// TIA Portal V20 export
Screen "170FX1Layout"  1276x673
  ScreenItem "Graphic view_1" at 215,132 size 858x332  Type=HmiGraphicView
  ScreenItem "Line_Header_X0_Y64" at 0,64 size 1276x0  Type=HmiLine
  ScreenItem "permanentareaborderrectangle" at 0,0 size 0x0  Type=HmiRectangle
  ScreenItem "Button_Back" at 2,2 size 90x60  Type=HmiButton
  ScreenItem "Move_Legend" at 1182,2 size 90x60  Type=HmiButton
  ScreenItem "Fusszeile_Button_ManualOPMode1_2" at 279,2 size 90x60  Type=HmiButton
  ScreenItem "文本域_3" at 1107,71 size 139x22  Type=HmiTextBox
  ScreenItem "LSicar_Valve8Pos_LeftHomeRightWork_WithPB_5" at 1099,95 size 160x53  Type=HmiFaceplateContainer
  ScreenItem "文本域_1" at 1107,160 size 156x23  Type=HmiTextBox
  ScreenItem "LSicar_Valve8Pos_LeftHomeRightWork_WithPB_1" at 1099,183 size 160x53  Type=HmiFaceplateContainer
  ScreenItem "文本域_22" at 1124,475 size 104x23  Type=HmiTextBox
  ScreenItem "面板容器_23" at 1171,508 size 96x32  Type=HmiFaceplateContainer
  ScreenItem "面板容器_22" at 1061,508 size 96x32  Type=HmiFaceplateContainer
  ScreenItem "面板容器_2" at 1087,4 size 88x58  Type=HmiFaceplateContainer
  ScreenItem "OPMode1_Blocked" at 1164,6 size 14x14  Type=HmiGraphicView
  ScreenItem "OPMode4_Foreground_Blocked" at 1088,4 size 88x58  Type=HmiGraphicView
  ScreenItem "Fusszeile_Button_ManualOPMode1_1" at 95,2 size 90x60  Type=HmiButton
  ScreenItem "面板容器_1" at 57,315 size 58x46  Type=HmiFaceplateContainer
  ScreenItem "面板容器_10" at 308,579 size 153x58  Type=HmiFaceplateContainer
  ScreenItem "Line_2" at 294,129 size 134x113  Type=HmiLine
  ScreenItem "面板容器_5" at 428,138 size 143x50  Type=HmiFaceplateContainer
  ScreenItem "Fusszeile_Button_ManualOPMode1_3" at 187,2 size 90x60  Type=HmiButton
  ScreenItem "文本域_6" at 428,97 size 140x40  Type=HmiTextBox
  ScreenItem "文本域_8" at 31,272 size 100x40  Type=HmiTextBox
  ScreenItem "文本域_13" at 313,557 size 140x20  Type=HmiTextBox
  ScreenItem "文本域_14" at 936,-172 size 140x40  Type=HmiTextBox
  ScreenItem "Title_ScreenOverview_X390_Y2_1" at 384,5 size 510x57  Type=HmiTextBox
  ScreenItem "文本域_26" at 907,541 size 140x40  Type=HmiTextBox
  ScreenItem "面板容器_15" at 910,583 size 149x54  Type=HmiFaceplateContainer
  ScreenItem "Line_19" at 989,402 size 32x137  Type=HmiLine
  ScreenItem "Line_1" at 443,402 size 106x106  Type=HmiLine
  ScreenItem "Line_3" at 302,399 size 75x157  Type=HmiLine
  ScreenItem "面板容器_4" at 492,529 size 153x58  Type=HmiFaceplateContainer
  ScreenItem "文本域_2" at 497,507 size 140x20  Type=HmiTextBox
  ScreenItem "面板容器_3" at 28,207 size 143x50  Type=HmiFaceplateContainer
  ScreenItem "文本域_4" at 28,166 size 140x40  Type=HmiTextBox
  ScreenItem "文本域_7" at 17,392 size 140x40  Type=HmiTextBox
  ScreenItem "面板容器_6" at 17,433 size 143x50  Type=HmiFaceplateContainer
  ScreenItem "Line_4" at 169,190 size 106x107  Type=HmiLine
  ScreenItem "Line_5" at 159,353 size 112x60  Type=HmiLine
  ScreenItem "Line_6" at 248,168 size 12x107  Type=HmiLine
  ScreenItem "面板容器_7" at 215,122 size 143x50  Type=HmiFaceplateContainer
  ScreenItem "文本域_9" at 215,81 size 140x40  Type=HmiTextBox
  ScreenItem "Line_7" at 171,371 size 89x165  Type=HmiLine
  ScreenItem "面板容器_8" at 83,577 size 143x50  Type=HmiFaceplateContainer
  ScreenItem "文本域_10" at 83,536 size 140x40  Type=HmiTextBox
  ScreenItem "Line_8" at 134,297 size 185x23  Type=HmiLine
  ScreenItem "Line_9" at 437,186 size 225x134  Type=HmiLine
  ScreenItem "面板容器_9" at 662,148 size 58x46  Type=HmiFaceplateContainer
  ScreenItem "文本域_11" at 636,105 size 100x40  Type=HmiTextBox
  ScreenItem "文本域_27" at 6,114 size 120x40  Type=HmiTextBox
  ScreenItem "文本域_5" at 5,69 size 120x40  Type=HmiTextBox
